SUBAPPLICATION OPC_TO_AR2_OUT (* Remote-Wert per OPC-UA als AR2 + AR-Spiegel VALUE_OUT (ohne VT) *)
  (* Standard: 61499-2; Description: Copyright (c) 2026 Meisterschulen am Ostbahnhof This program and the accompanying materials are made available under the terms of the Eclipse Public License 2.0 which is available at https://www.eclipse.org/legal/epl-2.0/ SPDX-License-Identifier: EPL-2.0 *)
  (* Version 1.0, 2026-10-28, Franz Höpfinger, Meisterschulen am Ostbahnhof, Kopie von MyLib::sys::NumericValue_TO_AR2_OPC ohne NumericValue_PHYSA/Q_NumericValue_PHYSA/AR_LAST_2, fuer Stationen ohne VT (keine isobus_UT-Libs). Wie MyLib::sys::OPC_TO_AR2, aber mit VALUE_OUT. *)
  PACKAGE MyLib::sys;
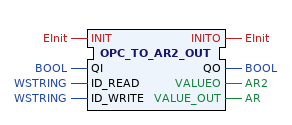
  EVENT_INPUT
    INIT : EInit; (* Initialization Request *)
  END_EVENT
  EVENT_OUTPUT
    INITO : EInit; (* Initialization Confirm *)
  END_EVENT
  VAR_INPUT
    QI : BOOL := TRUE; (* Quality Input - TRUE to enable service *)
    ID_READ : WSTRING; (* Remote-Subscribe-Adresse (REAL, ACTION=SUBSCRIBE) *)
    ID_WRITE : WSTRING; (* Remote-Echo-Adresse (REAL, ACTION=PUBLISH) *)
  END_VAR
  VAR_OUTPUT
    QO : BOOL; (* Quality Output - TRUE if service executed successfully *)
  END_VAR
  PLUGS
    VALUEO : adapter::types::bidirectional::AR2;
    VALUE_OUT : adapter::types::unidirectional::AR; (* AR-Spiegel des aktuellen Werts (= AR_TO_AR2.AR_OUT) *)
  END_PLUGS
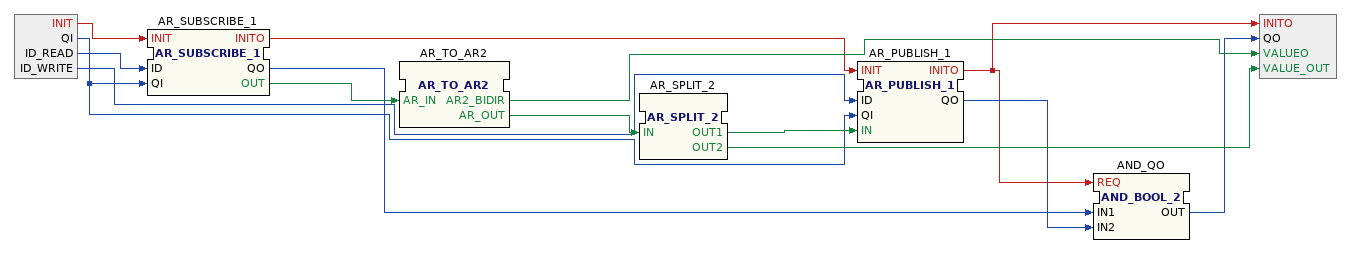
  FBS
    AR_SUBSCRIBE_1 : adapter::net::AR_SUBSCRIBE_1;
    AR_TO_AR2 : adapter::conversion::bidirectional::AR_TO_AR2;
    AR_SPLIT_2 : adapter::events::unidirectional::AR_SPLIT_2;
    AR_PUBLISH_1 : adapter::net::AR_PUBLISH_1;
    AND_QO : iec61131::booleanOperators::AND_BOOL_2;
  END_FBS
  EVENT_CONNECTIONS
    INIT TO AR_SUBSCRIBE_1.INIT;
    AR_SUBSCRIBE_1.INITO TO AR_PUBLISH_1.INIT;
    AR_PUBLISH_1.INITO TO INITO;
    AR_PUBLISH_1.INITO TO AND_QO.REQ;
  END_CONNECTIONS
  DATA_CONNECTIONS
    ID_READ TO AR_SUBSCRIBE_1.ID;
    ID_WRITE TO AR_PUBLISH_1.ID;
    QI TO AR_SUBSCRIBE_1.QI;
    QI TO AR_PUBLISH_1.QI;
    AR_SUBSCRIBE_1.QO TO AND_QO.IN1;
    AR_PUBLISH_1.QO TO AND_QO.IN2;
    AND_QO.OUT TO QO;
  END_CONNECTIONS
  ADAPTER_CONNECTIONS
    AR_SUBSCRIBE_1.OUT TO AR_TO_AR2.AR_IN;
    AR_TO_AR2.AR2_BIDIR TO VALUEO;
    AR_TO_AR2.AR_OUT TO AR_SPLIT_2.IN;
    AR_SPLIT_2.OUT1 TO AR_PUBLISH_1.IN;
    AR_SPLIT_2.OUT2 TO VALUE_OUT;
  END_CONNECTIONS
END_SUBAPPLICATION
